(* CODESYS project Energy.export

Project tree, tasks and I/O mapping:
  visualisation Energy
*)

// /Energy
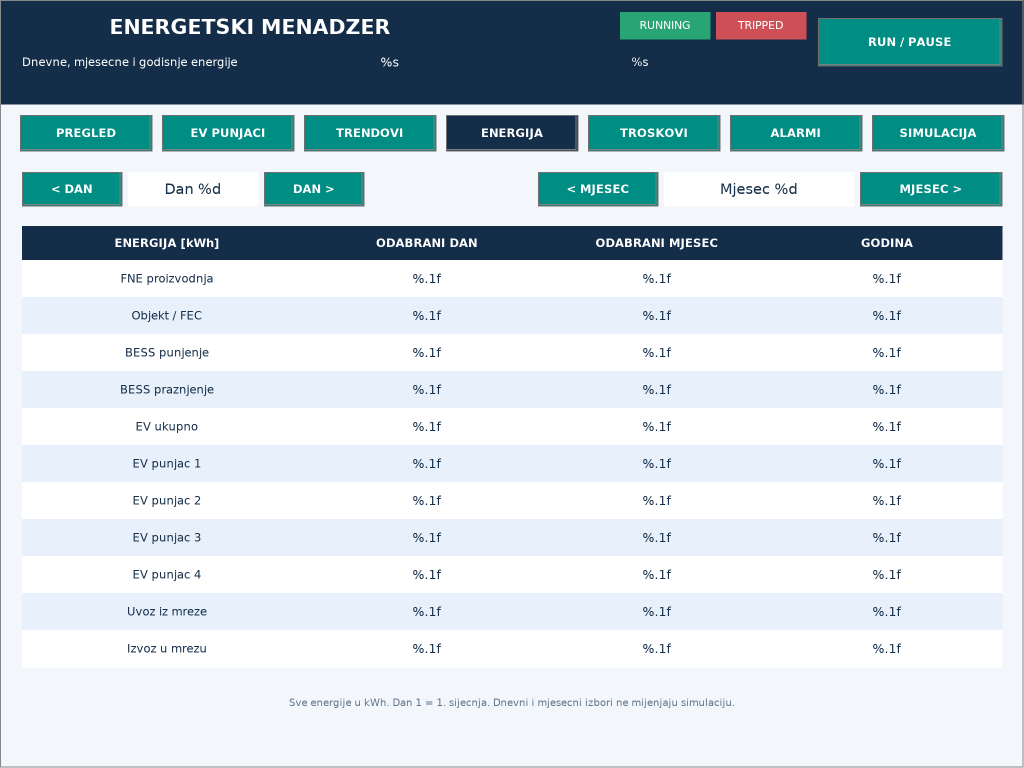
VISUALIZATION Energy  // 1024x768
    Rectangle (0,0 1024x768)
    Rectangle (0,0 1024x104)
    Rectangle (20,10 460x34), "ENERGETSKI MENADZER"
    Rectangle (20,48 220x28), "Dnevne, mjesecne i godisnje energije"
    Rectangle (260,49 260x26), "%s", text variable: Team_HMI.sDateTime
    Rectangle (530,49 220x26), "%s", text variable: Team_HMI.sPriceMode
    Button (818,18 184x48), "RUN / PAUSE"
        toggle SimCtrl.run
    Rectangle (620,12 90x27), "PAUSED", invisible if: SimCtrl.run
    Rectangle (620,12 90x27), "RUNNING", invisible if: NOT SimCtrl.run
    Rectangle (716,12 90x27), "TRIPPED", invisible if: NOT SimCtrl.tripped
    Button (20,115 132x36), "PREGLED"
        OnMouseClick:  Assign=Overview, Type=Assignment
    Button (162,115 132x36), "EV PUNJACI"
        OnMouseClick:  Assign=EVs, Type=Assignment
    Button (304,115 132x36), "TRENDOVI"
        OnMouseClick:  Assign=Trends, Type=Assignment
    Button (446,115 132x36), "ENERGIJA"
        OnMouseClick:  Assign=Energy, Type=Assignment
    Button (588,115 132x36), "TROSKOVI"
        OnMouseClick:  Assign=Costs, Type=Assignment
    Button (730,115 132x36), "ALARMI"
        OnMouseClick:  Assign=Alarms, Type=Assignment
    Button (872,115 132x36), "SIMULACIJA"
        OnMouseClick:  Assign=Controls, Type=Assignment
    Button (22,172 100x34), "< DAN"
        OnMouseClick: execute { Team_HMI.iSelDay := MAX(0, Team_HMI.iSelDay - 1); }
    Rectangle (128,172 130x34), "Dan %d", text variable: Team_HMI.iSelDay + 1
    Button (264,172 100x34), "DAN >"
        OnMouseClick: execute { Team_HMI.iSelDay := MIN(364, Team_HMI.iSelDay + 1); }
    Button (538,172 120x34), "< MJESEC"
        OnMouseClick: execute { Team_HMI.iSelMonth := MAX(1, Team_HMI.iSelMonth - 1); }
    Rectangle (664,172 190x34), "Mjesec %d", text variable: Team_HMI.iSelMonth
    Button (860,172 142x34), "MJESEC >"
        OnMouseClick: execute { Team_HMI.iSelMonth := MIN(12, Team_HMI.iSelMonth + 1); }
    Rectangle (22,226 290x34), "ENERGIJA [kWh]"
    Rectangle (312,226 230x34), "ODABRANI DAN"
    Rectangle (542,226 230x34), "ODABRANI MJESEC"
    Rectangle (772,226 230x34), "GODINA"
    Rectangle (22,260 290x37), "FNE proizvodnja"
    Rectangle (312,260 230x37), "%.1f", text variable: Team_Log.aDay[Team_HMI.iSelDay].E_fne
    Rectangle (542,260 230x37), "%.1f", text variable: Team_Log.aMonth[Team_HMI.iSelMonth].E_fne
    Rectangle (772,260 230x37), "%.1f", text variable: Team_Results.E_fne
    Rectangle (22,297 290x37), "Objekt / FEC"
    Rectangle (312,297 230x37), "%.1f", text variable: Team_Log.aDay[Team_HMI.iSelDay].E_fec
    Rectangle (542,297 230x37), "%.1f", text variable: Team_Log.aMonth[Team_HMI.iSelMonth].E_fec
    Rectangle (772,297 230x37), "%.1f", text variable: Team_Results.E_fec
    Rectangle (22,334 290x37), "BESS punjenje"
    Rectangle (312,334 230x37), "%.1f", text variable: Team_Log.aDay[Team_HMI.iSelDay].E_bess_chg
    Rectangle (542,334 230x37), "%.1f", text variable: Team_Log.aMonth[Team_HMI.iSelMonth].E_bess_chg
    Rectangle (772,334 230x37), "%.1f", text variable: Team_Results.E_bess_chg
    Rectangle (22,371 290x37), "BESS praznjenje"
    Rectangle (312,371 230x37), "%.1f", text variable: Team_Log.aDay[Team_HMI.iSelDay].E_bess_dch
    Rectangle (542,371 230x37), "%.1f", text variable: Team_Log.aMonth[Team_HMI.iSelMonth].E_bess_dch
    Rectangle (772,371 230x37), "%.1f", text variable: Team_Results.E_bess_dch
    Rectangle (22,408 290x37), "EV ukupno"
    Rectangle (312,408 230x37), "%.1f", text variable: Team_Log.aDay[Team_HMI.iSelDay].E_ev
    Rectangle (542,408 230x37), "%.1f", text variable: Team_Log.aMonth[Team_HMI.iSelMonth].E_ev
    Rectangle (772,408 230x37), "%.1f", text variable: Team_Results.E_ev
    Rectangle (22,445 290x37), "EV punjac 1"
    Rectangle (312,445 230x37), "%.1f", text variable: Team_Log.aDay[Team_HMI.iSelDay].E_ev_ch[0]
    Rectangle (542,445 230x37), "%.1f", text variable: Team_Log.aMonth[Team_HMI.iSelMonth].E_ev_ch[0]
    Rectangle (772,445 230x37), "%.1f", text variable: Team_Results.E_ev_ch[0]
    Rectangle (22,482 290x37), "EV punjac 2"
    Rectangle (312,482 230x37), "%.1f", text variable: Team_Log.aDay[Team_HMI.iSelDay].E_ev_ch[1]
    Rectangle (542,482 230x37), "%.1f", text variable: Team_Log.aMonth[Team_HMI.iSelMonth].E_ev_ch[1]
    Rectangle (772,482 230x37), "%.1f", text variable: Team_Results.E_ev_ch[1]
    Rectangle (22,519 290x37), "EV punjac 3"
    Rectangle (312,519 230x37), "%.1f", text variable: Team_Log.aDay[Team_HMI.iSelDay].E_ev_ch[2]
    Rectangle (542,519 230x37), "%.1f", text variable: Team_Log.aMonth[Team_HMI.iSelMonth].E_ev_ch[2]
    Rectangle (772,519 230x37), "%.1f", text variable: Team_Results.E_ev_ch[2]
    Rectangle (22,556 290x37), "EV punjac 4"
    Rectangle (312,556 230x37), "%.1f", text variable: Team_Log.aDay[Team_HMI.iSelDay].E_ev_ch[3]
    Rectangle (542,556 230x37), "%.1f", text variable: Team_Log.aMonth[Team_HMI.iSelMonth].E_ev_ch[3]
    Rectangle (772,556 230x37), "%.1f", text variable: Team_Results.E_ev_ch[3]
    Rectangle (22,593 290x37), "Uvoz iz mreze"
    Rectangle (312,593 230x37), "%.1f", text variable: Team_Log.aDay[Team_HMI.iSelDay].E_import
    Rectangle (542,593 230x37), "%.1f", text variable: Team_Log.aMonth[Team_HMI.iSelMonth].E_import
    Rectangle (772,593 230x37), "%.1f", text variable: Team_Results.E_import
    Rectangle (22,630 290x37), "Izvoz u mrezu"
    Rectangle (312,630 230x37), "%.1f", text variable: Team_Log.aDay[Team_HMI.iSelDay].E_export
    Rectangle (542,630 230x37), "%.1f", text variable: Team_Log.aMonth[Team_HMI.iSelMonth].E_export
    Rectangle (772,630 230x37), "%.1f", text variable: Team_Results.E_export
    Rectangle (22,689 980x27), "Sve energije u kWh. Dan 1 = 1. sijecnja. Dnevni i mjesecni izbori ne mijenjaju simulaciju."
END_VISUALIZATION
